(* IEC 61131-3 sources: JingjiangArm/moonboxpro_arm_8.4/Application/Application/任务列表/TensionTask/张力控制/收放料/张力调整, 5 files *)

(* ---- KS_ThisStepThatByStraightLine.st ---- *)
(*@CES
Name=KS_ThisStepThatByStraightLine
Type=FunctionBlock
TypeGuid=6f9dac99-8de1-4efc-8465-68ac443b7d08
Guid=7e0684ca-8029-4adc-9883-37fc94a520b5
HasDeclaration=True
HasImplementation=True
*)
{DECLARATION}
FUNCTION KS_ThisStepThatByStraightLine : BOOL(*到达目标值标志*)
VAR_INPUT
	i_rThis:REAL;(*起始值 用于计算变化量*)
	i_rThat:REAL;(*目标值*)
	i_prCur:POINTER TO REAL;(*当前值*)
	i_iStepTime:INT:=10;(*S*)
	i_iCycleTime:INT:=20;(*程序执行时间*)
	i_xFlag_Cut_end:BOOL;
END_VAR
VAR
	rDel: REAL;
	rCur: REAL;
END_VAR
{IMPLEMENTATION}
IF i_iStepTime=0 THEN
	i_iStepTime:=10*1000;
ELSE
	i_iStepTime:=i_iStepTime*1000;
END_IF(*ms即10s*)

rDel:=(i_rThat-i_rThis)/i_iStepTime*i_iCycleTime;(*计算变化量*)
rDel:=ABS(rDel);

IF i_prCur<>0 THEN
(*有个小bug 目标值从a切到b未到达b的时候又切到a可能会存在不变化的问题；
针对该问题 我们将变化量值切换为固定值|2019.4.11.095538*)

	IF rDel=0 AND i_prCur^<>i_rThat THEN
		rDel:=ABS(10.0/i_iStepTime*i_iCycleTime);(*固定变化量*)
	END_IF

	IF i_xFlag_Cut_end THEN
		i_prCur^:=i_rThat;
	ELSE
		IF i_prCur^>i_rThat THEN
			i_prCur^:=i_prCur^-rDel;
			IF i_prCur^<i_rThat THEN
				i_prCur^:=i_rThat;
			END_IF
		ELSIF i_prCur^<i_rThat THEN
			i_prCur^:=i_prCur^+rDel;
			IF i_prCur^>i_rThat THEN
				i_prCur^:=i_rThat;
			END_IF
		ELSE
			i_prCur^:=i_rThat;
		END_IF
	END_IF

	IF i_prCur^=i_rThat THEN
		KS_ThisStepThatByStraightLine:=TRUE;
	END_IF
ELSE
	RETURN;
END_IF

(* ---- KS_FB_Exchange.st ---- *)
(*@CES
Name=KS_FB_Exchange
Type=FunctionBlock
TypeGuid=6f9dac99-8de1-4efc-8465-68ac443b7d08
Guid=72852f5d-8de1-4e86-9ad2-e4d3bdb444a6
HasDeclaration=True
HasImplementation=True
*)
{DECLARATION}
FUNCTION_BLOCK KS_FB_Exchange
VAR_INPUT
	i_xCut_end: BOOL;
END_VAR
VAR_OUTPUT
END_VAR
VAR
	lrPreDia: LREAL;
	lrVel_Temp: LREAL;
	PI: LREAL:=3.1415926;
	xParamExchanged: BOOL;
END_VAR
VAR_IN_OUT
	io_rDiam_Cur: REAL;(*当前卷径*)
	io_rDiam_New: REAL;(*新卷径，单位是mm*)
	io_rVel_UwRw: REAL;(* 当前速度*)
	io_rVel_PreDrv: REAL;(*预驱速度*)

END_VAR
{IMPLEMENTATION}
(*该功能块在裁切换料完成之后进行预驱以及当前轴的卷径切换*
*同时要放在收放料裁切换料标志清零之前 *)(*当前速度的单位是R/MIN 预驱的速度单位是M/MIN*)

IF i_xCut_end AND NOT xParamExchanged THEN(*裁切完成后进行卷径，速度切换*)

	lrVel_Temp:=io_rVel_UwRw*io_rDiam_Cur*PI/1000;	(*将输入的当前速度转换为预驱速度 M/MIN*)
	io_rVel_UwRw:=io_rVel_PreDrv/io_rDiam_New/PI*1000;(*将预驱线速度转换为角速度R/MIN赋值给当前速度*)
	io_rVel_PreDrv:=lrVel_Temp;

(*将新卷径值赋给当前卷径值，将当前卷径值赋给新卷径值*)
	lrPreDia:=io_rDiam_Cur;
	io_rDiam_Cur:=io_rDiam_New;
	io_rDiam_New:=lrPreDia;
	xParamExchanged:=TRUE;
ELSIF NOT i_xCut_end THEN
	lrPreDia:=io_rDiam_New;
	xParamExchanged:=FALSE;
END_IF

(* ---- KS_FB_GetKpid.st ---- *)
(*@CES
Name=KS_FB_GetKpid
Type=FunctionBlock
TypeGuid=6f9dac99-8de1-4efc-8465-68ac443b7d08
Guid=b21071f8-c6ec-480a-ba8e-e12362a853f5
HasDeclaration=True
HasImplementation=True
*)
{DECLARATION}
FUNCTION_BLOCK KS_FB_GetKpid
VAR_INPUT
	i_xEn: BOOL;
	i_xCutFinish: BOOL;(*裁切完成标志*)
	i_iCycleTime_Plc: INT;(*周期时间*)
	i_rInitP: REAL;(*初始PID*)
	i_rInitI: REAL;
	i_rInitD: REAL;
	i_rDia_Cur: REAL;(*当前料卷卷径*)
	i_rThresholdCoeff: REAL:= 0.1;(*阈值系数*)
	i_xFlag_Cut_End: BOOL;
	i_xCutDneResetPidEn						: BOOL := FALSE;
	i_piCutDneResetPidMultiple				: POINTER TO INT;(*接料后放料PID放大倍数|单位修改为%2019.11.26.074236*)
	i_iCutDneResetPidRemainTime				: INT;(*保持时间S*)
	i_iCutDneResetPidToDefaultTime			: INT;(*恢复到默认的时间*)

	i_xSmallDiaMulEn						: BOOL:= FALSE;
	i_iSmallDiaMulSa						: INT:=200;(*进入该方式的启动卷径|大卷径*)
	i_iSmallDiaMulEd						: INT:=100;(*结束的卷径|写死为最小卷径*)
	i_iSmallDiaMulSa_Coeff					: INT:=100;(*系数|单位%*)
	i_iSmallDiaMulEd_Coeff					: INT:=300;(*系数|单位%*)
	i_xPseudoRandomTsting					: BOOL;(*伪随机测试标志||PID使用默认值*)
END_VAR
VAR_OUTPUT
	o_xEno									: BOOL;(*Indicated to i_xEn|*)
	o_iErNo									: INT;(*错误代码\-1:参数错误|*)
	o_rKp									: REAL;(*实际要使用的Kp*)
	o_rKi									: REAL;(*实际要使用的Ki*)
	o_rKd									: REAL;(*实际要使用的Kd*)
END_VAR
VAR
	iDiaStep								: INT;(*卷径区间步进*)
	iDia_Min								: INT:=200;(*卷径区间小*)
	iDia_Max								: INT:=2000;(*卷径区间大*)
	iMaxNum									: INT;
	aiDiaInterval							: ARRAY [0..30] OF INT;(*卷径区间数组*)
	iN										: INT;
	axArea									: ARRAY [1..31] OF BOOL;
	rInitDia								: REAL;
	xInit									: BOOL;
	iCurArea								: INT;
	iMinDia									: INT;
	iMaxDia									: INT;
	rMinDiaThreshold						: REAL;
	rMaxDiaThreshold						: REAL;
	xPreCutFinsh							: BOOL;
	rAverageDia							: REAL;
	arPid									: ARRAY [1..3] OF REAL;(*当前的pid*)
	arPrePid								: ARRAY [1..3] OF REAL;(*之前的pid*)
	axDne									: ARRAY [1..3] OF BOOL;(*变化完成*)
	fbKS_FB_GetPIDMul						: KS_FB_GetPIDMul;
	rCutDneResetPidMul						: REAL;
	rSmallDia_Coeff							: REAL;
END_VAR

{IMPLEMENTATION}
o_xEno:= i_xEn;
o_iErNo:= 0;

IF i_xEn THEN
	iDiaStep:=100;(*分段区间的间隔*)
	iMaxNum:=(iDia_Max-iDia_Min)/iDiaStep+1;
	aiDiaInterval[0]:=90;(*取一个较小的卷径值*)(*最后的区间为90，200，300，400，500。。。2000*)
	FOR iN:=1 TO iMaxNum-1 BY 1 DO
		aiDiaInterval[iN]:=iDia_Min+iDiaStep*(iN-1);
	END_FOR
	aiDiaInterval[iMaxNum]:=iDia_Max;
	(*以小中卷径的中间值作为和初始pid对应的卷径大小*)
	rInitDia:=350;
	IF i_rDia_Cur>iDia_Max THEN(*最大输入卷径*)
		i_rDia_Cur:=iDia_Max;
	END_IF

	IF i_rDia_Cur<90 THEN(*最小输入卷径*)
		i_rDia_Cur:=90;
	END_IF

	FOR iN:=1 TO 30 BY  1 DO(*清除标志*)
		axArea[iN]:=FALSE;
	END_FOR
	IF i_rDia_Cur<=aiDiaInterval[1] THEN(*小于最小卷径的时候*)
		axArea[1]:=TRUE;
	ELSE
		FOR iN:=1 TO iMaxNum-1 BY 1 DO
			IF i_rDia_Cur>aiDiaInterval[iN] AND  i_rDia_Cur<=aiDiaInterval[iN+1] THEN
				axArea[iN+1]:=TRUE;
				EXIT;
			END_IF
		END_FOR
	END_IF

	FOR iN:=1 TO iMaxNum BY  1 DO(*定位上个周期卷径所在的区间*)
		IF axArea[iN] THEN
			IF NOT xInit THEN
				xInit:=TRUE;
				iCurArea:=iN;
			END_IF
			IF iCurArea>iN THEN(*卷径值从大区间变为小区间*)
				iMinDia:=aiDiaInterval[iN-1];
				iMaxDia:=aiDiaInterval[iN];
				rMinDiaThreshold:=0;
				rMaxDiaThreshold:=iMaxDia*i_rThresholdCoeff;
			ELSIF  iCurArea<iN THEN(*卷径值从大区间变为小区间*)
				iMinDia:=aiDiaInterval[iN-1];
				iMaxDia:=aiDiaInterval[iN];
				rMinDiaThreshold:=iMinDia*i_rThresholdCoeff;
				rMaxDiaThreshold:=0;
			ELSE
				iMinDia:=aiDiaInterval[iN-1];
				iMaxDia:=aiDiaInterval[iN];
				rMinDiaThreshold:=0;
				rMaxDiaThreshold:=0;
			END_IF

			IF rMaxDiaThreshold>iDiaStep/2 THEN
				rMaxDiaThreshold:=iDiaStep/2;
			END_IF

			IF rMinDiaThreshold>iDiaStep/2 THEN
				rMinDiaThreshold:=iDiaStep/2;
			END_IF
			EXIT;
		END_IF
	END_FOR
	IF i_xCutFinish AND NOT xPreCutFinsh THEN(*裁切换料完成了*)(*裁切换料完成时不再考虑阈值问题2018.9.6.210051添加by liu.yt*)
		rMinDiaThreshold:=0;
		rMaxDiaThreshold:=0;
	END_IF
	xPreCutFinsh:=i_xCutFinish;

	IF (i_rDia_Cur>(iMinDia+rMinDiaThreshold)) AND (i_rDia_Cur<=(iMaxDia-rMaxDiaThreshold)) THEN
		iCurArea:=iN;
	END_IF

	IF iCurArea>iN THEN
		iCurArea:=iN+1;
		IF iCurArea>iMaxNum THEN
			iCurArea:=iMaxNum;
		END_IF
	ELSIF  iCurArea<iN THEN
		iCurArea:=iN-1;
		IF iCurArea<1 THEN
			iCurArea:=1;
		END_IF
	ELSE;
	END_IF

	iMinDia:=aiDiaInterval[iCurArea-1];
	iMaxDia:=aiDiaInterval[iCurArea];
	rAverageDia:=INT_TO_REAL(iMinDia+iMaxDia)/2;
	IF rAverageDia<>0 THEN
		arPid[1]:=i_rInitP*rInitDia/rAverageDia;
		arPid[2]:=i_rInitI*rInitDia/rAverageDia;
		arPid[3]:=i_rInitD*rInitDia/rAverageDia;
	ELSE
		arPid[1]:=i_rInitP;
		arPid[2]:=i_rInitI;
		arPid[3]:=i_rInitD;
		o_iErNo:=o_iErNo+1;
	END_IF

	(*--------------------------------------------------|2019.11.28.152830_*)
	(*裁切换料PID放大功能|小卷径pid增大倍数|*)
	fbKS_FB_GetPIDMul(
		i_xEn:= TRUE,
		i_xCutFinish:= i_xCutFinish,
		i_xCutDneResetPidEn:= i_xCutDneResetPidEn,
		i_piCutDneResetPidMultiple:= i_piCutDneResetPidMultiple,
		i_iCutDneResetPidRemainTime:= i_iCutDneResetPidRemainTime,
		i_iCutDneResetPidToDefaultTime:= i_iCutDneResetPidToDefaultTime,
		i_xSmallDiaMulEn:= i_xSmallDiaMulEn,
		i_rDia_Cur:= i_rDia_Cur,
		i_iSmallDiaMulSa:= i_iSmallDiaMulSa,
		i_iSmallDiaMulEd:= i_iSmallDiaMulEd,
		i_iSmallDiaMulSa_Coeff:= i_iSmallDiaMulSa_Coeff,
		i_iSmallDiaMulEd_Coeff:= i_iSmallDiaMulEd_Coeff,
		i_iCycleTime_Plc:= i_iCycleTime_Plc,
		o_xEn=> ,
		o_rCutDneResetPidMul=> rCutDneResetPidMul,
		o_rSmallDia_Coeff=> rSmallDia_Coeff);
	IF rCutDneResetPidMul<>1 THEN
		arPid[1]:=arPid[1]*rCutDneResetPidMul;
(*2022.9.13.100541*)
(*
		alrPid[2]:=alrPid[2]*rCutDneResetPidMul;
		alrPid[3]:=alrPid[3]*rCutDneResetPidMul;
*)
	ELSIF rSmallDia_Coeff<>1 THEN
		arPid[1]:=arPid[1]*rSmallDia_Coeff;
(*只放大了p值*)
(*
		alrPid[2]:=alrPid[2]*rSmallDia_Coeff;
		alrPid[3]:=alrPid[3]*rSmallDia_Coeff;
*)
	END_IF
	(*--------------------------------------------------|End|*)

(*2019.4.4.114213增加了pid切换直线变换逻辑|liu.yt*)
	IF NOT xInit THEN
		xInit:=TRUE;
		arPrePid:=arPid;
	END_IF
(**********************************)
(*2019.6.12.104845|niu.j|PID切换时间由10s改成5s，现场反馈裁切后摆臂震荡*)
	IF i_iCycleTime_Plc=0 THEN
		i_iCycleTime_Plc:= 20;
	END_IF
	axDne[1]:=KS_ThisStepThatByStraightLine(
								arPrePid[1],
								arPid[1],
								ADR(o_rKp),
								5,
								i_iCycleTime_Plc,
								i_xFlag_Cut_end);
	IF axDne[1] THEN
		arPrePid[1]:=arPid[1];
	END_IF
(*\\\\\\\\\\\\\\\\\\\\\\\\\\\\\\\\\*)
	axDne[2]:=KS_ThisStepThatByStraightLine(
								arPrePid[2],
								arPid[2],
								ADR(o_rKi),
								5,
								i_iCycleTime_Plc,
								i_xFlag_Cut_end);
	IF axDne[2] THEN
		arPrePid[2]:=arPid[2];
	END_IF
(*##################################*)
	axDne[3]:=KS_ThisStepThatByStraightLine(
								arPrePid[3],
								arPid[3],
								ADR(o_rKd),
								5,
								i_iCycleTime_Plc,
								i_xFlag_Cut_end);
	IF axDne[3] THEN
		arPrePid[3]:=arPid[3];
	END_IF
	(*2022.11.2.104544*)
	(*2022.9.10.101415 增加了伪随机的测试代码|2022.9.10.101424*)
	IF i_xPseudoRandomTsting THEN(*在处于伪随机测试|pid使用输入值*)
		o_rKp:=i_rInitP;
		o_rKi:=i_rInitI;
		o_rKd:=i_rInitD;
	END_IF

ELSE
	;
END_IF

(* ---- KS_FB_GetPIDMul.st ---- *)
(*@CES
Name=KS_FB_GetPIDMul
Type=FunctionBlock
TypeGuid=6f9dac99-8de1-4efc-8465-68ac443b7d08
Guid=0d44f791-d70b-4464-9f10-fe1428a728b2
HasDeclaration=True
HasImplementation=True
*)
{DECLARATION}
FUNCTION_BLOCK KS_FB_GetPIDMul
VAR_INPUT
	i_xEn:BOOL;
	i_xCutFinish:BOOL;(*裁切完成标志*)
	i_xCutDneResetPidEn:BOOL;
	i_piCutDneResetPidMultiple:POINTER TO INT;(*接料后放料PID放大倍数|单位修改为%2019.11.26.074236*)
	i_iCutDneResetPidRemainTime:INT;(*保持时间S*)
	i_iCutDneResetPidToDefaultTime:INT;(*恢复到默认的时间*)

	(*2019.11.22.084326  增加小卷径时pid放大一定倍数的逻辑|按照直线方式变化|大卷径小系数，小卷径大系数*)
	i_xSmallDiaMulEn:BOOL;
	i_rDia_Cur:LREAL;
	i_iSmallDiaMulSa:INT:=200;(*进入该方式的启动卷径|大卷径*)
	i_iSmallDiaMulEd:INT:=100;(*结束的卷径|写死为最小卷径*)
	i_iSmallDiaMulSa_Coeff:INT:=100;(*系数|单位%*)
	i_iSmallDiaMulEd_Coeff:INT:=300;(*系数|单位%*)
	i_iCycleTime_Plc: INT;(*周期时间*)
END_VAR
VAR_OUTPUT
	o_xEn:BOOL;
	o_rCutDneResetPidMul:REAL;(*接料后倍数|单位是1*)
	o_rSmallDia_Coeff: REAL;(*小卷径倍数|单位是%*)
END_VAR
VAR
	xCutDneCanResetPid: BOOL:=FALSE;(*可以放大pid标志*)
	xCutDneResetPidResume: BOOL:=FALSE;(*pid恢复标志*)
	iCutDneResetPidMaxMul:INT:=2;(*最大倍数*)
	lrCutDneResetPidMul: LREAL;
	iCnt: INT;

	(*小卷启动pid增大一定倍数逻辑使用的变量*)
	lrCoeff: LREAL;
	xCoeffEn: BOOL;
	lrK: LREAL;
END_VAR
{IMPLEMENTATION}
(*2019.10.12.212315 裁切完成后pid值增大一定的倍数功能*)
IF i_piCutDneResetPidMultiple<>0 THEN
	IF i_piCutDneResetPidMultiple^>1000 THEN(*倍数最大10倍  最小1倍*)
		 i_piCutDneResetPidMultiple^:=1000;
	ELSIF i_piCutDneResetPidMultiple^<=0 THEN
		i_piCutDneResetPidMultiple^:=100;
	END_IF
	iCutDneResetPidMaxMul:=i_piCutDneResetPidMultiple^;(*PID放大的最大倍数*)
ELSE
	iCutDneResetPidMaxMul:=100;
END_IF

IF i_xCutFinish AND NOT xCutDneCanResetPid THEN(*裁切完成*)
	xCutDneCanResetPid:=TRUE;
END_IF

IF i_iCycleTime_Plc=0 THEN
	i_iCycleTime_Plc:= 20;
END_IF
lrCutDneResetPidMul:=100;
IF i_xCutDneResetPidEn THEN
	IF xCutDneCanResetPid THEN
		lrCutDneResetPidMul:=INT_TO_LREAL(iCutDneResetPidMaxMul);
		iCnt:=iCnt+1;
		IF iCnt>=i_iCutDneResetPidRemainTime*1000/i_iCycleTime_Plc THEN(*持续时间.若为0则从最大倍数开始递减*)
			xCutDneCanResetPid:=FALSE;
			xCutDneResetPidResume:=TRUE;
			iCnt:=0;
		END_IF
	ELSE
		IF xCutDneResetPidResume THEN
			IF iCnt>=i_iCutDneResetPidToDefaultTime*1000/i_iCycleTime_Plc THEN
				xCutDneResetPidResume:=FALSE;
			ELSE
				iCnt:=iCnt+1;
				IF i_iCutDneResetPidToDefaultTime<>0 THEN
					lrCutDneResetPidMul:=INT_TO_LREAL(iCutDneResetPidMaxMul)-
						INT_TO_LREAL(iCutDneResetPidMaxMul-100)/
						i_iCutDneResetPidToDefaultTime/1000*i_iCycleTime_Plc*iCnt;
				END_IF
			END_IF
		ELSE
			iCnt:=0;
		END_IF
	END_IF
ELSE
	xCutDneCanResetPid:=FALSE;
	xCutDneResetPidResume:=FALSE;
	iCnt:=0;
END_IF
o_rCutDneResetPidMul:=LREAL_TO_REAL(lrCutDneResetPidMul/100);
IF lrCutDneResetPidMul=100 THEN o_rCutDneResetPidMul:=1;END_IF

(*2019.10.7.093811 在小卷径的时候针对pid增加了系数|200直径--->100直径|Liu.yt*)
IF i_rDia_Cur<=i_iSmallDiaMulSa THEN
	xCoeffEn:=TRUE;
ELSIF i_rDia_Cur>=i_iSmallDiaMulSa+20 THEN(*增加了浮动区间20mm*)
	xCoeffEn:=FALSE;
END_IF

IF i_xSmallDiaMulEn THEN;
ELSE
	xCoeffEn:=FALSE;
END_IF

IF xCoeffEn THEN
	IF i_iSmallDiaMulEd<>i_iSmallDiaMulSa THEN(*起始和结束的卷径不相等*)
		(*2023.2.17.151740*)
		lrK:=INT_TO_LREAL(i_iSmallDiaMulEd_Coeff-i_iSmallDiaMulSa_Coeff)/(i_iSmallDiaMulEd-i_iSmallDiaMulSa);
	ELSE
		lrK:=0;(*卷径一样的时候 按照大卷径系数输出！*)
	END_IF

	lrCoeff:=lrK*i_rDia_Cur+(i_iSmallDiaMulSa_Coeff-lrK*i_iSmallDiaMulSa);
	IF lrCoeff>i_iSmallDiaMulEd_Coeff THEN lrCoeff:=i_iSmallDiaMulEd_Coeff;END_IF
	IF lrCoeff<i_iSmallDiaMulSa_Coeff THEN lrCoeff:=i_iSmallDiaMulSa_Coeff;END_IF
ELSE
	lrCoeff:=100;
END_IF
o_rSmallDia_Coeff:= LREAL_TO_REAL(lrCoeff/100.0);
IF lrCoeff=100 THEN o_rSmallDia_Coeff:=1;END_IF

(* ---- KS_FB_UwRw_TensionCTL.st ---- *)
(*@CES
Name=KS_FB_UwRw_TensionCTL
Type=FunctionBlock
TypeGuid=6f9dac99-8de1-4efc-8465-68ac443b7d08
Guid=db71b4fc-851f-434f-8f6c-f56559c6fd2e
HasDeclaration=True
HasImplementation=True
*)
{DECLARATION}
FUNCTION_BLOCK KS_FB_UwRw_TensionCTL
VAR_INPUT
	i_xEn: BOOL;
	i_xIsDebugMode:BOOL;(*调试模式*)
	i_xNegative_PiValue:BOOL;(*pi取反*)
	i_xMachineRev:BOOL;(*反向走料信号*)
	i_xCutPressed: BOOL;(*裁切压辊合压标志*)
	i_xCancelPWhenCut:BOOL;(*裁切输出时取消p值标志|延时恢复*)
	i_rVel_Film: REAL;(*料膜速度*)
	i_rAI: REAL;(*传感器反馈*)
	i_prVel_AxisCur: POINTER TO REAL;(*速度值-转速*)
	i_rKp: REAL;(*P值*)
	i_rKi: REAL;(*I值*)
	i_rKd: REAL;(*D值*)
	i_iCycleTime_Plc:INT;(*程序执行周期*)
	i_xAccDecingCompensateEn:BOOL;
	i_rFeedforwordValue_Uw: REAL;
	i_iCut_PIInput_Time: INT; (*放料裁切PI投入时间*)
	(*放料翻转架补偿转速值|2021.7.26.092528*)
	i_rDeltaW_RPMIN:REAL;
	(*2021.9.13.132503|放料接料补偿值|窄方波+微分*)
	i_rSpliceCompensate:REAL;
	(*2021.8.26.170700|增加收放料主转速变化量-和是否使用预估卷径相关|使用则有值-否则=0*)
	i_rMailVel:REAL;
	i_rDiamCurAxis:REAL;(*当前卷径*)

END_VAR
VAR_OUTPUT
	o_xEn: BOOL;
	o_iErNo: INT;
	o_rStep:REAL;
	o_rPi_Value:REAL;
	o_rTotalPiValue:REAL;(*总的pi控制量*)
END_VAR
VAR
	iN: INT;
	iSum: INT:=100;
	rSum: REAL;
	rAverage: REAL;
	rPreVel_Film : REAL;
	arAI_Sum: ARRAY [1..200] OF REAL:= [200(0)];
	rUwRwForward_Step: REAL;(*前馈值*)
	arPID: ARRAY [1..3] OF REAL;
	rCoeff_I_UwCut: REAL;(*2024.8.20.103518|裁切时积分系数 *)
	xFlag_CancleP: BOOL;(*取消P值标志*)
	iCut_PIInput_Count: INT:=0;(*放料裁切PID投入计时*)
	rPIValue: REAL;
	iNum_Old: INT:= 5;(*D值上个值的位置*)
END_VAR

{IMPLEMENTATION}
o_xEn:= i_xEn;
o_iErNo:= 0;
rSum:= 0;
FOR iN:= iSum TO 2 BY -1 DO(*滑窗的时候顺道算一下和*)
	arAI_Sum[iN]:= arAI_Sum[iN-1];
	rSum:= rSum+arAI_Sum[iN];
END_FOR
arAI_Sum[1]:= i_rAI;
rSum:= rSum+arAI_Sum[1];
rAverage:= rSum/iSum;(*计算平均值*)
arPID[1]:= i_rKp;
arPID[2]:= i_rKi;
arPID[3]:= i_rKd;

IF i_xEn THEN
	IF i_prVel_AxisCur<>0 AND i_rVel_Film>0 THEN
		(*先计算前馈值*)
		rUwRwForward_Step:= 0;
		IF i_xAccDecingCompensateEn THEN(*料膜加速完成了，才使用前馈*)
			IF i_rVel_Film<>rPreVel_Film AND rPreVel_Film<>0 AND i_rVel_Film>=10 THEN
				rUwRwForward_Step:= (i_rVel_Film-rPreVel_Film)/rPreVel_Film*i_prVel_AxisCur^*
								BOOL_TO_INT(i_xAccDecingCompensateEn);
			ELSE
				;
			END_IF
		END_IF

		(*小卷高速前馈*)
		IF i_rAI<0 THEN(*如果放料变松了，我们就不再需要这种前馈补偿了*)
			i_rFeedforwordValue_Uw:= 0;
		END_IF
		rUwRwForward_Step:= rUwRwForward_Step+ i_rFeedforwordValue_Uw;
		(*2024.8.22.093024 增加了放料裁切后积分的系数随摆臂位置的变化*)
		(*2024.8.20.103438 在接料的时候积分逐步加大-根据摆臂位置*)
		IF ABS(i_rAI)>2 THEN
			rCoeff_I_UwCut:=1.0/5.0;
		ELSIF ABS(i_rAI)>1 THEN
			rCoeff_I_UwCut:=1.0/4.0;
		ELSIF ABS(i_rAI)>0.5 THEN
			rCoeff_I_UwCut:=1.0/3.0;
		ELSE
			rCoeff_I_UwCut:=1.0/2.0;
		END_IF
		IF i_xCancelPWhenCut THEN
			xFlag_CancleP:= TRUE;
			iCut_PIInput_Count:= 0;
			i_rKp:= i_rKp*rCoeff_I_UwCut;
		ELSE
			IF xFlag_CancleP THEN
				IF i_iCut_PIInput_Time<= i_iCycleTime_Plc*iCut_PIInput_Count THEN(*PI投入时间到了*)
					iCut_PIInput_Count:=0;
					xFlag_CancleP:=FALSE;
				ELSE
					iCut_PIInput_Count:= iCut_PIInput_Count+1;
					i_rKp:= i_rKp*rCoeff_I_UwCut;
				END_IF
			END_IF
		END_IF
		rPIValue:= LREAL_TO_REAL(i_rKp/1000*i_rAI+
			i_rKd/100*(arAI_Sum[1]-arAI_Sum[iNum_Old]));
		IF i_xCutPressed THEN (*主要是放料*)
			rPIValue:=0;
		END_IF
		IF i_xNegative_PiValue THEN(*PI取反|*)
			rPIValue:=-rPIValue;
		END_IF

		IF i_xMachineRev THEN(*反向走料|只需要取反调整量-主速度会在输出部分取反*)
			rPIValue:=-rPIValue;
		END_IF
		(*2021.7.26.092414 增加了翻转架运动补偿转速|*)
		IF i_prVel_AxisCur^+rPIValue+rUwRwForward_Step+i_rDeltaW_RPMIN+i_rMailVel+i_rSpliceCompensate<0 THEN
			i_prVel_AxisCur^:=0;
		ELSE
			i_prVel_AxisCur^:=i_prVel_AxisCur^+rPIValue+rUwRwForward_Step+i_rDeltaW_RPMIN+i_rMailVel+i_rSpliceCompensate;
			o_rTotalPiValue:=o_rTotalPiValue+rPIValue;(*统计pi控制量@2023.09.09.120357*)
		END_IF
		IF i_xIsDebugMode THEN
			IF i_rDiamCurAxis<>0 THEN
				i_prVel_AxisCur^:= LREAL_TO_REAL(i_rVel_Film*1000.0/gc_lrPi/i_rDiamCurAxis);
			END_IF
		END_IF
		o_rPi_Value:= rPIValue;
		o_rStep:= rUwRwForward_Step;
		o_xEn:= TRUE;
	ELSE(*非印刷状态，料膜速度=0*)
		FOR iN:=1 TO iSum BY 1 DO
			arAI_Sum[iN]:=0;
		END_FOR
		iCut_PIInput_Count:=0;
		xFlag_CancleP:=FALSE;
		o_rPi_Value:= 0;
		o_rStep:= 0;
		o_xEn:= FALSE;
	END_IF
	rPreVel_Film:= i_rVel_Film;
ELSE
	;
END_IF
